Staubli VAL3: teachPoint.pgx

program teachPoint(num x_nIndex)
  local bool l_bResult
  local tool l_tTool
begin
  link(l_tTool,flange)
//  call savedata:getTool(1,l_tTool)
  l_bResult=userPageConfirm("是否记录点位："+toString("",x_nIndex)+"?")
  if l_bResult
    safeTemp:sSPoint[x_nIndex].pPointRx=here(flange,world)
    safeTemp:libSave()
    delay(0.1)
  endIf
end
